Fanuc KAREL source: kb00131.KL

PROGRAM KB00131
%STACKSIZE=65535
%PRIORITY=65535
%NOLOCKGROUP
VAR
P1 : STRING[80]
P2 : BOOLEAN
P3 : INTEGER
P4 : INTEGER
P5 : STRING[80]
P6 : INTEGER
P7 : INTEGER
BEGIN
P1='A'
P2=TRUE
P3=1
P4=1
P5='A'
P6=1
P7=1
PIPE_CONFIG(P1,P2,P3,P4,P5,P6,P7)
END KB00131
